SUBAPPLICATION SubApp_PC_B (* Geraet B: Adder (opcua.adoc): SUBSCRIBE Num1/Num2 -> F_ADD -> PUBLISH Result, Werte z.B. per UaExpert *)
  (* Standard: 61499-2; Description: Copyright (c) 2026 Meisterschulen am Ostbahnhof This program and the accompanying materials are made available under the terms of the Eclipse Public License 2.0 which is available at https://www.eclipse.org/legal/epl-2.0/ SPDX-License-Identifier: EPL-2.0 *)
  (* Version 1.0, 2026-10-18, Franz Höpfinger, Meisterschulen am Ostbahnhof, opcua.adoc-Beispiel auf zwei Geraeten *)
  PACKAGE subapp::Training_14_OPC_UA_RES;
  IMPORT VV::const::OPC_UA::myOpcUaAddresses::T14_NUM1_READ;
  IMPORT VV::const::OPC_UA::myOpcUaAddresses::T14_NUM2_READ;
  IMPORT VV::const::OPC_UA::myOpcUaAddresses::T14_RESULT_WRITE;
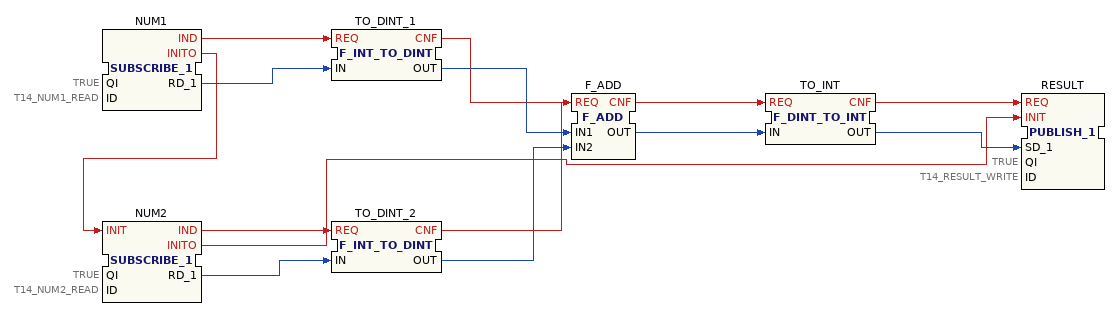
  FBS
    NUM1 : iec61499::net::SUBSCRIBE_1(QI := TRUE, ID := T14_NUM1_READ);
    NUM2 : iec61499::net::SUBSCRIBE_1(QI := TRUE, ID := T14_NUM2_READ);
    TO_DINT_1 : iec61131::conversion::F_INT_TO_DINT;
    TO_DINT_2 : iec61131::conversion::F_INT_TO_DINT;
    F_ADD : iec61131::arithmetic::F_ADD;
    TO_INT : iec61131::conversion::F_DINT_TO_INT;
    RESULT : iec61499::net::PUBLISH_1(QI := TRUE, ID := T14_RESULT_WRITE);
  END_FBS
  EVENT_CONNECTIONS
    NUM1.IND TO TO_DINT_1.REQ;
    NUM2.IND TO TO_DINT_2.REQ;
    TO_DINT_1.CNF TO F_ADD.REQ;
    TO_DINT_2.CNF TO F_ADD.REQ;
    F_ADD.CNF TO TO_INT.REQ;
    TO_INT.CNF TO RESULT.REQ;
    NUM1.INITO TO NUM2.INIT;
    NUM2.INITO TO RESULT.INIT;
  END_CONNECTIONS
  DATA_CONNECTIONS
    NUM1.RD_1 TO TO_DINT_1.IN;
    NUM2.RD_1 TO TO_DINT_2.IN;
    TO_DINT_1.OUT TO F_ADD.IN1;
    TO_DINT_2.OUT TO F_ADD.IN2;
    F_ADD.OUT TO TO_INT.IN;
    TO_INT.OUT TO RESULT.SD_1;
  END_CONNECTIONS
END_SUBAPPLICATION
